(* IEC 61131-3 sources: 2026_Projet_YGO_ExcavatriceDragage/CODE/J_SUPERVISION (part 3) *)

(* ---- FB_TroubleshootingView.st ---- *)
(* ═══════════════════════════════════════════════════════════════
   🕵️♂️ FB_TroubleshootingView — Mise en forme lecture seule pour dépannage
   ───────────────────────────────────────────────────────────────
   📄 Doc : DOC/AF/AF_Partie-14_Fonction_Troubleshooting/FB_TroubleshootingView_v1.2.md
   🔗 Producteur unique de GVL_Troubleshooting.* — instancié UNE SEULE FOIS,
      dans PRG_07_Supervision, après §3 Projections IHM.
   🔒 Lecture seule stricte : aucune VAR_OUTPUT de commande, aucun calcul métier,
      aucune fusion de source — pure recopie de faits déjà publiés ailleurs.
   ⚠️ WinchM2 est typé ST_WinchBenneHMI (pas ST_WinchHMI comme WinchM1) : ce lot
      (LOT_TROUBLESHOOTING_VIEW_ET_WINCHHMI) a introduit ST_WinchBenneHMI pour porter
      Bucket côté M2 uniquement (GVL_IHM.M2TreuilBenne) — adaptation du port fiche §3
      nécessaire suite à AC5 (Bucket retiré de ST_WinchHMI commun M1/M2).
   Écriture GVL directe : seule exception au principe "pas de GVL comme bus de
      commande" (AF_Partie-03 §5) — GVL_Troubleshooting n'est jamais relue par un FB
      métier, uniquement par Watch CODESYS / export SCADA dépannage (fiche §3/§7).
   ⚠️ Idx201_JoystickSelected (ContexteMachineGlobal) lit GVL_IHM.Modes.Cmd.TglJoystickMaster
      directement (variable globale IEC 61131-3, visible sans passage par VAR_INPUT) — ce
      port n'est pas dans la table fiche §3 mais le producteur exact est documenté fiche §5.1.
   ═══════════════════════════════════════════════════════════════ *)
FUNCTION_BLOCK PUBLIC FB_TroubleshootingView
VAR_INPUT
    Enable                   : BOOL; (* --> [CMD] TRUE en permanence — fiche §3, aucune condition de scan *)

    (* 📡 PRG_02_Acquisition *)
    HwIn                     : ST_HardwareImage;   (* --> [HW] Image entrées qualifiées *)
    HwReal                   : ST_HardwareImage;   (* --> [HW] Image entrées réelles *)
    InputModuleFault         : BOOL;   (* --> [HW] Défaut module d'entrée *)
    LocalDigitalIoOk         : BOOL; (* --> [HW] Mirroir Network.InputModules — pas de champ ST_Chain* dédié ce lot *)
    Vh0800EndOk              : BOOL; (* --> [HW] idem *)
    Vh0808EtpOk              : BOOL; (* --> [HW] idem *)

    (* 🎚️ PRG_03_Modes_Cycle *)
    Auth                     : ST_Modes_Autorisations;   (* --> [SAFE] Autorisations machine *)

    (* 🛗 PRG_04_Treuils_Benne — demandes publiques déjà arbitrées *)
    M1LogicRequestSpeedCmd_Pct : REAL;   (* --> [CMD] Consigne vitesse M1 *)
    M1LogicRequestDirection    : INT;   (* --> [CMD] Sens M1 *)
    M2LogicRequestSpeedCmd_Pct : REAL;   (* --> [CMD] Consigne vitesse M2 *)
    M2LogicRequestDirection    : INT;   (* --> [CMD] Sens M2 *)
    WinchBothMotionDirection : INT;   (* --> [CMD] Direction couplée *)
    WinchBothMotionActive    : BOOL;   (* --> [CMD] Demande couplée active *)
    CycleAutoBusy                : BOOL;   (* --> [HW] Cycle auto actif *)
    CycleM1SpeedTgt_Pct          : REAL;   (* --> [CMD] Consigne cycle M1 *)
    CycleM2SpeedTgt_Pct          : REAL;   (* --> [CMD] Consigne cycle M2 *)
    CycleBucketOpen              : BOOL;   (* --> [HW] Benne ouverte cycle *)
    CycleTargetPosition          : INT;   (* --> [CMD] Cible cycle *)

    (* 🎭 GVL_Simulation *)
    SimulationModeActive     : BOOL;   (* --> [TST] Mode simulation *)
    SimWinchActive           : BOOL;   (* --> [TST] Sim treuils *)
    SimTranslationActive     : BOOL;   (* --> [TST] Sim translation *)
    SimOperatorActive        : BOOL;   (* --> [TST] Sim opérateur *)
    SimSafetyActive          : BOOL;   (* --> [TST] Sim sécurité *)

    (* 🛗 GVL_IHM — images publiques déjà produites *)
    WinchM1                  : ST_WinchHMI;      (* --> [HW] GVL_IHM.M1TreuilRetenue *)
    WinchM2                  : ST_WinchBenneHMI; (* --> [HW] GVL_IHM.M2TreuilBenne — porte Bucket *)
    Sync                     : ST_SyncHMI;       (* --> [HW] GVL_IHM.M1M2Sync *)
    Translation              : ST_TranslationHMI;(* --> [HW] GVL_IHM.M3Translation *)
    Commun                   : ST_CommunHMI;     (* --> [HW] GVL_IHM.Commun *)
    Network                  : ST_NetworkDiagHMI;(* --> [HW] GVL_IHM.Network *)
    JoystickHMI              : ST_JoystickHMI;   (* --> [HW] GVL_IHM.JOY1Joystick *)
    Permits                  : ST_PermitVisibilityHMI; (* --> [DIAG] Vue unique des permis produite par PRG_07 *)

    (* 🛡️ Sorties publiques AU produites par PRG_06_Outputs *)
    EmergencyState           : ST_Safety_Emergency_State;   (* --> [SAFE] État AU *)
    EmergencyDiag            : ST_Safety_Emergency_Diag;   (* --> [SAFE] Diagnostic AU *)
    PowerCutOffActive        : BOOL;   (* --> [SAFE] Coupure puissance *)
    ArmingPulseActive        : BOOL;   (* --> [SAFE] Impulsion réarmement *)
    MaintainAActive          : BOOL;   (* --> [SAFE] Maintien canal A *)
    MaintainBActive          : BOOL;   (* --> [SAFE] Maintien canal B *)

    (* 📤 Ordres finaux produits par PRG_06_Outputs, après barrière et protecteurs *)
    Outputs                  : ST_OutputsInterPrg; (* --> [CMD] Ordres actionneurs finaux *)
    CmdM3DriveFreqWord       : WORD;   (* --> [CMD] Consigne finale variateur M3 [0.01 Hz] *)

    (* 🔄 Séquenceur de cycle semi-automatique *)
    CycleReady               : BOOL;   (* --> [STAT] Séquenceur prêt *)
    CycleDone                : BOOL;   (* --> [STAT] Séquenceur terminé *)
    CycleError               : BOOL;   (* --> [STAT] Séquenceur en erreur *)
    CycleErrorId             : WORD;   (* --> [DIAG] Code erreur séquenceur *)
    CycleFaultLatched        : BOOL;   (* --> [STAT] Défaut latché séquenceur (bloque AX0->AX1, exige Reset) *)
    CycleFaultLatchedId      : WORD;   (* --> [DIAG] Bitfield défaut latché figé *)
    CycleChecksInhibited     : BOOL;   (* --> [TST] Contrôles procédé inhibés *)
    CycleIgnoredCheckId      : WORD;   (* --> [DIAG] Contrôles procédé ignorés *)
    CycleForceStepResult     : STRING(120); (* --> [DIAG] Motif de rejet de la consigne de forcage de step (T358) *)
    CycleStep                : E_AutoCycleStep; (* --> [STAT] Étape courante *)
    CycleStepStr             : STRING(80);  (* --> [STAT] Libellé étape *)
    CycleStepAtError         : E_AutoCycleStep; (* --> [DIAG] Étape au défaut *)
    CycleWaitingForOperator  : BOOL;        (* --> [STAT] Attente action humaine *)
    CycleWaitingForProcess   : BOOL;        (* --> [STAT] Attente condition procédé *)
    CycleOperatorActionId    : WORD;        (* --> [DIAG] ID action attendue *)
    CycleOperatorAction      : STRING(120); (* --> [DIAG] Consigne explicite *)
    CycleExpectedAxis        : E_OperatorAxis; (* --> [STAT] Organe attendu *)
    CycleExpectedDirection   : INT;         (* --> [STAT] Sens attendu (-1, 0, +1) *)
    CycleStartRequest        : BOOL;   (* --> [CMD] Demande Start *)
    CycleAbortRequest        : BOOL;   (* --> [CMD] Demande Abort *)
    CycleTargetDepth_M       : REAL;   (* --> [CFG] Profondeur consigne *)
    CycleKoboldBottomTouch   : BOOL;   (* --> [HW] Contact fond *)
    CycleSpeedMismatchActive : BOOL;   (* --> [DIAG] Écart vitesse M1/M2 *)
    CycleLimitLegalReached   : BOOL;   (* --> [SAFE] Limite légale atteinte *)
    CycleWinchSyncError      : BOOL;   (* --> [SAFE] Erreur synchro treuils *)
    CycleM1SpeedStepApplied  : INT;    (* --> [HW] Palier vitesse appliqué M1 (0..5, causes 8/9 FB_CycleSemiAuto) *)
    CycleM2SpeedStepApplied  : INT;    (* --> [HW] Palier vitesse appliqué M2 (0..5, causes 8/9 FB_CycleSemiAuto) *)
    CycleAutoDiveM2Step5Active : BOOL; (* --> [STAT] Essai T291-A actif (M2 cible palier 5 en plongée) *)
    CycleM1SpeedStepAtFault  : INT;    (* --> [DIAG] Palier M1 appliqué, figé au moment du défaut (0..5) *)
    CycleM2SpeedStepAtFault  : INT;    (* --> [DIAG] Palier M2 appliqué, figé au moment du défaut (0..5) *)
    JoystickDeadmanArmed     : BOOL;   (* --> [CMD] Homme-mort armé *)
    JoystickAtNeutral        : BOOL;   (* --> [HW] Joystick au neutre *)
    HomedM1                  : BOOL;   (* --> [HW] Codeur M1 référencé *)
    HomedM2                  : BOOL;   (* --> [HW] Codeur M2 référencé *)

    (* 📐 Config effective limite haute — source _CommunCfgPersist (≠ copie IHM) *)
    CfgTopLimitM             : REAL;   (* --> [CFG] Limite haute active (m) = CfgCableLimitAscent_M *)

    (* 🕵️ PRG_04/05 — Trace de blocage terrain (cause priorisée + horodatage, produite
       par PRG_04 §8bis / PRG_05 §4bis, publiée via Data ; pure recopie ici) *)
    WinchM1Trace             : ST_TraceWinch;       (* --> [DIAG] Trace blocage treuil M1 *)
    WinchM2Trace             : ST_TraceWinch;       (* --> [DIAG] Trace blocage treuil M2 *)
    TranslationTrace         : ST_TraceTranslation; (* --> [DIAG] Trace blocage translation M3 *)
    MachineHoming            : ST_MachineHoming;    (* --> [DIAG] Etat public du cycle de homing conjoint *)
END_VAR
VAR_OUTPUT
    Ready                    : BOOL; (* <-- [STAT] Diagnostic interne minimal — fiche §3 *)
END_VAR

// 🛑 GATE — neutralisation ; aucune écriture GVL_Troubleshooting si Enable=FALSE
IF NOT Enable THEN
    Ready := FALSE;
    RETURN;
END_IF;
Ready := TRUE;

{region "§0 Contexte machine global"}
// === 🌐 0. ContexteMachineGlobal : ST_ChainContextGlobal (fiche §5.1) ===
GVL_Troubleshooting.A_ContexteMachineGlobal.Idx101_ModeActive        := Auth.Mode;
GVL_Troubleshooting.A_ContexteMachineGlobal.Idx102_SimulationEnabled := SimulationModeActive;
GVL_Troubleshooting.A_ContexteMachineGlobal.Idx103_JoystickCommOk    := Network.Joystick.Operational;
GVL_Troubleshooting.A_ContexteMachineGlobal.Idx201_JoystickSelected  := GVL_IHM.Modes.Cmd.TglJoystickMaster;
GVL_Troubleshooting.A_ContexteMachineGlobal.Idx202_BypassNetworkGlobal := Network.Bypass.Global;
GVL_Troubleshooting.A_ContexteMachineGlobal.Idx203_BypassSensorsGlobal := FALSE; // TBD non câblé - voir fiche §6 (agrégat multi-domaine à définir)
GVL_Troubleshooting.A_ContexteMachineGlobal.Idx301_EmergencyChainClosed := HwIn.Machine.EmergencyChainClosed_DI;
GVL_Troubleshooting.A_ContexteMachineGlobal.Idx302_PowerContactorEngaged := HwIn.Machine.PowerContactorEngaged_DI;
// Agrégat simple OR de faits déjà publiés (fiche §5.1) — pas un nouveau calcul métier
GVL_Troubleshooting.A_ContexteMachineGlobal.Idx303_SafeStopActiveAny := WinchM1.Safety.SafeStop OR WinchM2.Safety.SafeStop OR Translation.Safety.SafeStop;
GVL_Troubleshooting.A_ContexteMachineGlobal.Idx304_PowerCutOffActiveAny := WinchM1.Safety.PowerCutOff OR WinchM2.Safety.PowerCutOff OR Translation.Safety.PowerCutOff;
GVL_Troubleshooting.A_ContexteMachineGlobal.Idx401_HmiHeartbeatOk    := Commun.HeartbeatIhmOk;
GVL_Troubleshooting.A_ContexteMachineGlobal.Idx402_CycleAutoBusy     := CycleAutoBusy;

{endregion}

{region "§1 Levage synchronise M1/M2"}
// === 🛗 1. LevageSynchroniseM1M2 : ST_ChainWinchSync (fiche §5.2) ===
GVL_Troubleshooting.H_LevageSynchroniseM1M2.Idx101_M1_CablePos_M  := WinchM1.State.Position_M;
GVL_Troubleshooting.H_LevageSynchroniseM1M2.Idx102_M2_CablePos_M  := WinchM2.State.Position_M;
GVL_Troubleshooting.H_LevageSynchroniseM1M2.Idx103_SyncDelta_M    := Sync.State.DeltaPos_M;
GVL_Troubleshooting.H_LevageSynchroniseM1M2.Idx202_SyncEnabled_IHM := Sync.Cmd.SelSyncEnable;
GVL_Troubleshooting.H_LevageSynchroniseM1M2.Idx301_EmergencyChainClosed := HwIn.Machine.EmergencyChainClosed_DI;
GVL_Troubleshooting.H_LevageSynchroniseM1M2.Idx302_SyncFaultActive := Sync.State.Error;
GVL_Troubleshooting.H_LevageSynchroniseM1M2.Idx303_M1_AscentPermit := WinchM1.Safety.AscentPermit;
GVL_Troubleshooting.H_LevageSynchroniseM1M2.Idx304_M2_AscentPermit := WinchM2.Safety.AscentPermit;
GVL_Troubleshooting.H_LevageSynchroniseM1M2.Idx501_M1_CmdRelayFwd_DQ := Outputs.M1RelayFwd;
GVL_Troubleshooting.H_LevageSynchroniseM1M2.Idx502_M2_CmdRelayFwd_DQ := Outputs.M2RelayFwd;
// Idx201_JoyYRaw_Pct / Idx203_ArbitratedSpeed_Pct / Idx303-304_AscentPermit / Idx401_SyncMotionAllowed /
// Idx402-403_SetpointSpeed : non câblés — fiche §5.2 "(reste) champs à revoir un par un", laissés à
// leur valeur d'initialisation, pas de calcul inventé (fiche §7).

{endregion}

{region "§2 Levage unitaire M1/M2"}
// === 🛗 2. LevageUnitaireM1 / LevageUnitaireM2 : ST_ChainWinch (fiche §5.3) ===
// --- M1 ---
GVL_Troubleshooting.I_LevageUnitaireM1.Inputs_100.Idx101_EncoderRawPos := UDINT_TO_DINT(HwIn.Winch.COD1_PosValue);
GVL_Troubleshooting.I_LevageUnitaireM1.Inputs_100.Idx102_CablePos_M := WinchM1.State.Position_M;
GVL_Troubleshooting.I_LevageUnitaireM1.Inputs_100.Idx103_ContactorsReleased_DI := HwIn.Winch.M1_ContactorsReleased_DI;
GVL_Troubleshooting.I_LevageUnitaireM1.Inputs_100.Idx104_BrakeApplied := NOT HwIn.Winch.M1_BrakeIsOpen_DI;
GVL_Troubleshooting.I_LevageUnitaireM1.Inputs_100.Idx105_ThermalOk_DI := HwIn.Winch.M1_ThermalOk_DI;

GVL_Troubleshooting.I_LevageUnitaireM1.Demandes_200.Idx201_JoyRawPhysical_ANA := HwIn.Operator.JoyYRaw_ANA2;
GVL_Troubleshooting.I_LevageUnitaireM1.Demandes_200.Idx202_JoyScaledPhysical_Pct := JoystickHMI.State.AxisCmdY.Deflection;
GVL_Troubleshooting.I_LevageUnitaireM1.Demandes_200.Idx203_HmiManualCmd_BtnAscent := WinchM1.Cmd.BtnAscent;
GVL_Troubleshooting.I_LevageUnitaireM1.Demandes_200.Idx204_HmiManualCmd_BtnDescent := WinchM1.Cmd.BtnDescent;
GVL_Troubleshooting.I_LevageUnitaireM1.Demandes_200.Idx205_CycleAutoCmd_Pct := CycleM1SpeedTgt_Pct;
GVL_Troubleshooting.I_LevageUnitaireM1.Demandes_200.Idx206_ModeActive := Auth.Mode;
GVL_Troubleshooting.I_LevageUnitaireM1.Demandes_200.Idx207_BypassOperatorComm := WinchM1.Bypass.OperatorComm;
GVL_Troubleshooting.I_LevageUnitaireM1.Demandes_200.Idx208_ArbitratedSpeed_Pct := M1LogicRequestSpeedCmd_Pct;
GVL_Troubleshooting.I_LevageUnitaireM1.Demandes_200.Idx209_ArbitratedDirection := M1LogicRequestDirection;
GVL_Troubleshooting.I_LevageUnitaireM1.Demandes_200.Idx210_CoupledUserRequestDirection := WinchBothMotionDirection;
GVL_Troubleshooting.I_LevageUnitaireM1.Demandes_200.Idx211_CoupledUserRequestActive := WinchBothMotionActive;

GVL_Troubleshooting.I_LevageUnitaireM1.Safety_300.Idx301_EmergencyChainClosed := HwIn.Machine.EmergencyChainClosed_DI;
GVL_Troubleshooting.I_LevageUnitaireM1.Safety_300.Idx302_SafeStopActive := WinchM1.Safety.SafeStop;
GVL_Troubleshooting.I_LevageUnitaireM1.Safety_300.Idx303_PowerCutOffActive := WinchM1.Safety.PowerCutOff;
GVL_Troubleshooting.I_LevageUnitaireM1.Safety_300.Idx304_TopSensorPhysical_DI := HwIn.Winch.M1M2_TopPositionFree_DI;
GVL_Troubleshooting.I_LevageUnitaireM1.Safety_300.Idx305_TopSensorBypassActive := Commun.SimTopSensorBypassActive;
GVL_Troubleshooting.I_LevageUnitaireM1.Safety_300.Idx306_AscentPermitEffective := WinchM1.Safety.AscentPermit;
GVL_Troubleshooting.I_LevageUnitaireM1.Safety_300.Idx307_SlackCablePhysical_DI := NOT HwIn.Winch.M2_TensionedCable_DI; // Capteur unique partagé, même signal que SlackCableDetected M1
GVL_Troubleshooting.I_LevageUnitaireM1.Safety_300.Idx308_SlackCableBypassActive := Commun.SimSlackCableBypassActive;
GVL_Troubleshooting.I_LevageUnitaireM1.Safety_300.Idx309_DescendPermitEffective := WinchM1.Safety.DescendPermit;
GVL_Troubleshooting.I_LevageUnitaireM1.Safety_300.Idx310_ErrorOperatorComm := WinchM1.Safety.ErrorOperatorComm;
GVL_Troubleshooting.I_LevageUnitaireM1.Safety_300.Idx311_ErrorEncoder      := WinchM1.Safety.ErrorEncoder;
GVL_Troubleshooting.I_LevageUnitaireM1.Safety_300.Idx312_ErrorPhaseRotation:= WinchM1.Safety.ErrorPhaseRotation;
GVL_Troubleshooting.I_LevageUnitaireM1.Safety_300.Idx313_ErrorMecaA        := WinchM1.Safety.ErrorMecaA;
GVL_Troubleshooting.I_LevageUnitaireM1.Safety_300.Idx314_ErrorMecaB        := WinchM1.Safety.ErrorMecaB;
GVL_Troubleshooting.I_LevageUnitaireM1.Safety_300.Idx315_ErrorMecaC        := WinchM1.Safety.ErrorMecaC;
GVL_Troubleshooting.I_LevageUnitaireM1.Safety_300.Idx316_ErrorMecaD        := WinchM1.Safety.ErrorMecaD;
GVL_Troubleshooting.I_LevageUnitaireM1.Safety_300.Idx317_ErrorMecaE        := WinchM1.Safety.ErrorMecaE;
GVL_Troubleshooting.I_LevageUnitaireM1.Safety_300.Idx318_ErrorBrakeThermal := WinchM1.Safety.ErrorBrakeThermal;
GVL_Troubleshooting.I_LevageUnitaireM1.Safety_300.Idx319_ErrorOppositeDir  := WinchM1.Safety.ErrorOppositeDir;
GVL_Troubleshooting.I_LevageUnitaireM1.Safety_300.Idx320_ErrorNoMovement   := WinchM1.Safety.ErrorNoMovement;
// ⛔ Bloc "limite haute" — pourquoi la montée ne s'arrête pas (M1)
GVL_Troubleshooting.I_LevageUnitaireM1.Safety_300.Idx321_CfgTopLimitM               := CfgTopLimitM;
GVL_Troubleshooting.I_LevageUnitaireM1.Safety_300.Idx322_CablePosM                  := WinchM1.State.Position_M;
GVL_Troubleshooting.I_LevageUnitaireM1.Safety_300.Idx323_TopLimitReached            := WinchM1.Safety.CableLimitAscent;
GVL_Troubleshooting.I_LevageUnitaireM1.Safety_300.Idx324_AscentBlockedByTopLimit    := WinchM1.Safety.CableLimitAscent AND NOT (WinchM1.Bypass.TopLimitSoftware OR Commun.Bypass.TopLimitSoftware);
GVL_Troubleshooting.I_LevageUnitaireM1.Safety_300.Idx325_BypassTopLimitSoftware     := WinchM1.Bypass.TopLimitSoftware;
GVL_Troubleshooting.I_LevageUnitaireM1.Safety_300.Idx326_BypassTopLimitSoftCommun   := Commun.Bypass.TopLimitSoftware;
GVL_Troubleshooting.I_LevageUnitaireM1.Safety_300.Idx327_BypassTopLimitSwitch       := WinchM1.Bypass.TopLimitSwitch;
GVL_Troubleshooting.I_LevageUnitaireM1.Safety_300.Idx328_BypassTopLimitSwitchCommun := Commun.Bypass.TopLimitSwitch;
GVL_Troubleshooting.I_LevageUnitaireM1.Safety_300.Idx329_BypassGlobal               := WinchM1.Bypass.Global;
GVL_Troubleshooting.I_LevageUnitaireM1.Safety_300.Idx330_BypassGlobalCommun         := Commun.Bypass.Global;

GVL_Troubleshooting.I_LevageUnitaireM1.Control_400.Idx401_MotionAllowed := WinchM1.State.Ready;
GVL_Troubleshooting.I_LevageUnitaireM1.Control_400.Idx402_SpeedStepCalculated := WinchM1.State.StepNumber;
GVL_Troubleshooting.I_LevageUnitaireM1.Control_400.Idx403_SpeedRamp_Pct := WinchM1.State.SpeedCmd_Pct;
GVL_Troubleshooting.I_LevageUnitaireM1.Control_400.Idx404_BrakeReleaseAuthorized := WinchM1.State.BrakeCmd;
GVL_Troubleshooting.I_LevageUnitaireM1.Control_400.Idx405_FinalInterlockState := WinchM1.State.FinalInterlockState;
GVL_Troubleshooting.I_LevageUnitaireM1.Control_400.Idx406_FinalInterlockReason := WinchM1.State.FinalInterlockReason;
GVL_Troubleshooting.I_LevageUnitaireM1.Control_400.Idx407_FinalAuthorizedStep := WinchM1.State.FinalAuthorizedStep;
GVL_Troubleshooting.I_LevageUnitaireM1.Control_400.Idx408_BrakeCommandOpenConfirmed := WinchM1.State.BrakeCommandOpenConfirmed;
GVL_Troubleshooting.I_LevageUnitaireM1.Control_400.Idx409_BrakeTimeoutElapsed := WinchM1.State.FinalBrakeTimeoutElapsed;
GVL_Troubleshooting.I_LevageUnitaireM1.Control_400.Idx410_RestartDelayElapsed := WinchM1.State.FinalRestartDelayElapsed;
GVL_Troubleshooting.I_LevageUnitaireM1.Control_400.Idx411_StepDelayElapsed := WinchM1.State.FinalStepDelayElapsed;
GVL_Troubleshooting.I_LevageUnitaireM1.Control_400.Idx412_InTopSlowdownZone := WinchM1.State.InTopSlowdownZone;
GVL_Troubleshooting.I_LevageUnitaireM1.Control_400.Idx413_InBottomSlowdownZone := WinchM1.State.InBottomSlowdownZone;
GVL_Troubleshooting.I_LevageUnitaireM1.Control_400.Idx414_BottomLimitActiveM := WinchM1.State.BottomLimitActiveM;
GVL_Troubleshooting.I_LevageUnitaireM1.Control_400.Idx415_MotorRequest := WinchM1.State.FinalMotorRequest;
GVL_Troubleshooting.I_LevageUnitaireM1.Control_400.Idx416_RestartRequired := WinchM1.State.FinalRestartRequired;
GVL_Troubleshooting.I_LevageUnitaireM1.Control_400.Idx417_RestartInhibit := WinchM1.State.FinalRestartInhibit;
GVL_Troubleshooting.I_LevageUnitaireM1.Control_400.Idx418_NeutralRequestSeen := WinchM1.State.FinalNeutralRequestSeen;

GVL_Troubleshooting.I_LevageUnitaireM1.Outputs_500.Idx501_CmdRelayAscent_RQ := Outputs.M1RelayFwd;
GVL_Troubleshooting.I_LevageUnitaireM1.Outputs_500.Idx502_CmdRelayDescent_RQ := Outputs.M1RelayRev;
GVL_Troubleshooting.I_LevageUnitaireM1.Outputs_500.Idx503_CmdSpeedContactor1_DQ := Outputs.M1SpeedContactor1;
GVL_Troubleshooting.I_LevageUnitaireM1.Outputs_500.Idx504_CmdSpeedContactor4_DQ := Outputs.M1SpeedContactor4;
GVL_Troubleshooting.I_LevageUnitaireM1.Outputs_500.Idx505_CmdBrakeRelease_RQ := WinchM1.State.BrakeCmd;

// --- M2 (même patron, source WinchM2) ---
GVL_Troubleshooting.J_LevageUnitaireM2.Inputs_100.Idx101_EncoderRawPos := UDINT_TO_DINT(HwIn.Winch.COD2_PosValue);
GVL_Troubleshooting.J_LevageUnitaireM2.Inputs_100.Idx102_CablePos_M := WinchM2.State.Position_M;
GVL_Troubleshooting.J_LevageUnitaireM2.Inputs_100.Idx103_ContactorsReleased_DI := HwIn.Winch.M2_ContactorsReleased_DI;
GVL_Troubleshooting.J_LevageUnitaireM2.Inputs_100.Idx104_BrakeApplied := NOT HwIn.Winch.M2_BrakeIsOpen_DI;
GVL_Troubleshooting.J_LevageUnitaireM2.Inputs_100.Idx105_ThermalOk_DI := HwIn.Winch.M2_ThermalOk_DI;

GVL_Troubleshooting.J_LevageUnitaireM2.Demandes_200.Idx201_JoyRawPhysical_ANA := HwIn.Operator.JoyYRaw_ANA2;
GVL_Troubleshooting.J_LevageUnitaireM2.Demandes_200.Idx202_JoyScaledPhysical_Pct := JoystickHMI.State.AxisCmdY.Deflection;
GVL_Troubleshooting.J_LevageUnitaireM2.Demandes_200.Idx203_HmiManualCmd_BtnAscent := WinchM2.Cmd.BtnAscent;
GVL_Troubleshooting.J_LevageUnitaireM2.Demandes_200.Idx204_HmiManualCmd_BtnDescent := WinchM2.Cmd.BtnDescent;
GVL_Troubleshooting.J_LevageUnitaireM2.Demandes_200.Idx205_CycleAutoCmd_Pct := CycleM2SpeedTgt_Pct;
GVL_Troubleshooting.J_LevageUnitaireM2.Demandes_200.Idx206_ModeActive := Auth.Mode;
GVL_Troubleshooting.J_LevageUnitaireM2.Demandes_200.Idx207_BypassOperatorComm := WinchM2.Bypass.OperatorComm;
GVL_Troubleshooting.J_LevageUnitaireM2.Demandes_200.Idx208_ArbitratedSpeed_Pct := M2LogicRequestSpeedCmd_Pct;
GVL_Troubleshooting.J_LevageUnitaireM2.Demandes_200.Idx209_ArbitratedDirection := M2LogicRequestDirection;
GVL_Troubleshooting.J_LevageUnitaireM2.Demandes_200.Idx210_CoupledUserRequestDirection := WinchBothMotionDirection;
GVL_Troubleshooting.J_LevageUnitaireM2.Demandes_200.Idx211_CoupledUserRequestActive := WinchBothMotionActive;

GVL_Troubleshooting.J_LevageUnitaireM2.Safety_300.Idx301_EmergencyChainClosed := HwIn.Machine.EmergencyChainClosed_DI;
GVL_Troubleshooting.J_LevageUnitaireM2.Safety_300.Idx302_SafeStopActive := WinchM2.Safety.SafeStop;
GVL_Troubleshooting.J_LevageUnitaireM2.Safety_300.Idx303_PowerCutOffActive := WinchM2.Safety.PowerCutOff;
GVL_Troubleshooting.J_LevageUnitaireM2.Safety_300.Idx304_TopSensorPhysical_DI := HwIn.Winch.M1M2_TopPositionFree_DI;
GVL_Troubleshooting.J_LevageUnitaireM2.Safety_300.Idx305_TopSensorBypassActive := Commun.SimTopSensorBypassActive;
GVL_Troubleshooting.J_LevageUnitaireM2.Safety_300.Idx306_AscentPermitEffective := WinchM2.Safety.AscentPermit;
// Bug affichage MES 2026-09-04 : publiait TensionedCable_DI sans l'inverser -> cable
// tendu (bon) s'affichait comme "mou detecte". Logique securite reelle (PRG_04) deja
// correcte (NOT TensionedCable_DI) ; seul ce mirroir troubleshooting etait faux.
GVL_Troubleshooting.J_LevageUnitaireM2.Safety_300.Idx307_SlackCablePhysical_DI := NOT HwIn.Winch.M2_TensionedCable_DI;
GVL_Troubleshooting.J_LevageUnitaireM2.Safety_300.Idx308_SlackCableBypassActive := Commun.SimSlackCableBypassActive;
GVL_Troubleshooting.J_LevageUnitaireM2.Safety_300.Idx309_DescendPermitEffective := WinchM2.Safety.DescendPermit;
GVL_Troubleshooting.J_LevageUnitaireM2.Safety_300.Idx310_ErrorOperatorComm := WinchM2.Safety.ErrorOperatorComm;
GVL_Troubleshooting.J_LevageUnitaireM2.Safety_300.Idx311_ErrorEncoder      := WinchM2.Safety.ErrorEncoder;
GVL_Troubleshooting.J_LevageUnitaireM2.Safety_300.Idx312_ErrorPhaseRotation:= WinchM2.Safety.ErrorPhaseRotation;
GVL_Troubleshooting.J_LevageUnitaireM2.Safety_300.Idx313_ErrorMecaA        := WinchM2.Safety.ErrorMecaA;
GVL_Troubleshooting.J_LevageUnitaireM2.Safety_300.Idx314_ErrorMecaB        := WinchM2.Safety.ErrorMecaB;
GVL_Troubleshooting.J_LevageUnitaireM2.Safety_300.Idx315_ErrorMecaC        := WinchM2.Safety.ErrorMecaC;
GVL_Troubleshooting.J_LevageUnitaireM2.Safety_300.Idx316_ErrorMecaD        := WinchM2.Safety.ErrorMecaD;
GVL_Troubleshooting.J_LevageUnitaireM2.Safety_300.Idx317_ErrorMecaE        := WinchM2.Safety.ErrorMecaE;
GVL_Troubleshooting.J_LevageUnitaireM2.Safety_300.Idx318_ErrorBrakeThermal := WinchM2.Safety.ErrorBrakeThermal;
GVL_Troubleshooting.J_LevageUnitaireM2.Safety_300.Idx319_ErrorOppositeDir  := WinchM2.Safety.ErrorOppositeDir;
GVL_Troubleshooting.J_LevageUnitaireM2.Safety_300.Idx320_ErrorNoMovement   := WinchM2.Safety.ErrorNoMovement;
// ⛔ Bloc "limite haute" — pourquoi la montée ne s'arrête pas (M2, sans M2_LimitShift ici)
GVL_Troubleshooting.J_LevageUnitaireM2.Safety_300.Idx321_CfgTopLimitM               := CfgTopLimitM;
GVL_Troubleshooting.J_LevageUnitaireM2.Safety_300.Idx322_CablePosM                  := WinchM2.State.Position_M;
GVL_Troubleshooting.J_LevageUnitaireM2.Safety_300.Idx323_TopLimitReached            := WinchM2.Safety.CableLimitAscent;
GVL_Troubleshooting.J_LevageUnitaireM2.Safety_300.Idx324_AscentBlockedByTopLimit    := WinchM2.Safety.CableLimitAscent AND NOT (WinchM2.Bypass.TopLimitSoftware OR Commun.Bypass.TopLimitSoftware);
GVL_Troubleshooting.J_LevageUnitaireM2.Safety_300.Idx325_BypassTopLimitSoftware     := WinchM2.Bypass.TopLimitSoftware;
GVL_Troubleshooting.J_LevageUnitaireM2.Safety_300.Idx326_BypassTopLimitSoftCommun   := Commun.Bypass.TopLimitSoftware;
GVL_Troubleshooting.J_LevageUnitaireM2.Safety_300.Idx327_BypassTopLimitSwitch       := WinchM2.Bypass.TopLimitSwitch;
GVL_Troubleshooting.J_LevageUnitaireM2.Safety_300.Idx328_BypassTopLimitSwitchCommun := Commun.Bypass.TopLimitSwitch;
GVL_Troubleshooting.J_LevageUnitaireM2.Safety_300.Idx329_BypassGlobal               := WinchM2.Bypass.Global;
GVL_Troubleshooting.J_LevageUnitaireM2.Safety_300.Idx330_BypassGlobalCommun         := Commun.Bypass.Global;

GVL_Troubleshooting.J_LevageUnitaireM2.Control_400.Idx401_MotionAllowed := WinchM2.State.Ready;
GVL_Troubleshooting.J_LevageUnitaireM2.Control_400.Idx402_SpeedStepCalculated := WinchM2.State.StepNumber;
GVL_Troubleshooting.J_LevageUnitaireM2.Control_400.Idx403_SpeedRamp_Pct := WinchM2.State.SpeedCmd_Pct;
GVL_Troubleshooting.J_LevageUnitaireM2.Control_400.Idx404_BrakeReleaseAuthorized := WinchM2.State.BrakeCmd;
GVL_Troubleshooting.J_LevageUnitaireM2.Control_400.Idx405_FinalInterlockState := WinchM2.State.FinalInterlockState;
GVL_Troubleshooting.J_LevageUnitaireM2.Control_400.Idx406_FinalInterlockReason := WinchM2.State.FinalInterlockReason;
GVL_Troubleshooting.J_LevageUnitaireM2.Control_400.Idx407_FinalAuthorizedStep := WinchM2.State.FinalAuthorizedStep;
GVL_Troubleshooting.J_LevageUnitaireM2.Control_400.Idx408_BrakeCommandOpenConfirmed := WinchM2.State.BrakeCommandOpenConfirmed;
GVL_Troubleshooting.J_LevageUnitaireM2.Control_400.Idx409_BrakeTimeoutElapsed := WinchM2.State.FinalBrakeTimeoutElapsed;
GVL_Troubleshooting.J_LevageUnitaireM2.Control_400.Idx410_RestartDelayElapsed := WinchM2.State.FinalRestartDelayElapsed;
GVL_Troubleshooting.J_LevageUnitaireM2.Control_400.Idx411_StepDelayElapsed := WinchM2.State.FinalStepDelayElapsed;
GVL_Troubleshooting.J_LevageUnitaireM2.Control_400.Idx412_InTopSlowdownZone := WinchM2.State.InTopSlowdownZone;
GVL_Troubleshooting.J_LevageUnitaireM2.Control_400.Idx413_InBottomSlowdownZone := WinchM2.State.InBottomSlowdownZone;
GVL_Troubleshooting.J_LevageUnitaireM2.Control_400.Idx414_BottomLimitActiveM := WinchM2.State.BottomLimitActiveM;
GVL_Troubleshooting.J_LevageUnitaireM2.Control_400.Idx415_MotorRequest := WinchM2.State.FinalMotorRequest;
GVL_Troubleshooting.J_LevageUnitaireM2.Control_400.Idx416_RestartRequired := WinchM2.State.FinalRestartRequired;
GVL_Troubleshooting.J_LevageUnitaireM2.Control_400.Idx417_RestartInhibit := WinchM2.State.FinalRestartInhibit;
GVL_Troubleshooting.J_LevageUnitaireM2.Control_400.Idx418_NeutralRequestSeen := WinchM2.State.FinalNeutralRequestSeen;

GVL_Troubleshooting.J_LevageUnitaireM2.Outputs_500.Idx501_CmdRelayAscent_RQ := Outputs.M2RelayFwd;
GVL_Troubleshooting.J_LevageUnitaireM2.Outputs_500.Idx502_CmdRelayDescent_RQ := Outputs.M2RelayRev;
GVL_Troubleshooting.J_LevageUnitaireM2.Outputs_500.Idx503_CmdSpeedContactor1_DQ := Outputs.M2SpeedContactor1;
GVL_Troubleshooting.J_LevageUnitaireM2.Outputs_500.Idx504_CmdSpeedContactor4_DQ := Outputs.M2SpeedContactor4;
GVL_Troubleshooting.J_LevageUnitaireM2.Outputs_500.Idx505_CmdBrakeRelease_RQ := WinchM2.State.BrakeCmd;

{endregion}

{region "§3 Benne ouverture et fermeture"}
// === 🪣 3. BenneOuvertureFermeture : ST_ChainBucket (fiche §5.4, source WinchM2.Bucket) ===
GVL_Troubleshooting.K_BenneOuvertureFermeture.Idx101_BucketIsOpen := WinchM2.Bucket.State.MechState.IsOpen;
GVL_Troubleshooting.K_BenneOuvertureFermeture.Idx102_BucketIsClosed := WinchM2.Bucket.State.MechState.IsClosed;
GVL_Troubleshooting.K_BenneOuvertureFermeture.Idx103_OffsetPos_M := WinchM2.Bucket.State.ActiveOffset_M;
GVL_Troubleshooting.K_BenneOuvertureFermeture.Idx104_AutoSeqActive := WinchM2.Bucket.State.AutoBucketSeqActive;
GVL_Troubleshooting.K_BenneOuvertureFermeture.Idx105_StateIncoherent := WinchM2.Bucket.State.MechState.StateIncoherent;
GVL_Troubleshooting.K_BenneOuvertureFermeture.Idx106_FBState := WinchM2.Bucket.State.FBState;
GVL_Troubleshooting.K_BenneOuvertureFermeture.Idx107_LastPosM2Open_M := WinchM2.Bucket.State.MechState.LastPosM2Open;
GVL_Troubleshooting.K_BenneOuvertureFermeture.Idx108_LastPosM2Close_M := WinchM2.Bucket.State.MechState.LastPosM2Close;
GVL_Troubleshooting.K_BenneOuvertureFermeture.Idx109_BucketTooOpen := WinchM2.Bucket.State.MechState.TooOpen;
GVL_Troubleshooting.K_BenneOuvertureFermeture.Idx110_BucketTooClosed := WinchM2.Bucket.State.MechState.TooClosed;
GVL_Troubleshooting.K_BenneOuvertureFermeture.Idx111_BucketIsIntermediate := WinchM2.Bucket.State.MechState.IsIntermediate;
GVL_Troubleshooting.K_BenneOuvertureFermeture.Idx112_DeltaPosition_M := WinchM2.Bucket.State.DeltaPosition_M;
GVL_Troubleshooting.K_BenneOuvertureFermeture.Idx113_MachineHomed := WinchM2.Bucket.State.MachineHomed;
GVL_Troubleshooting.K_BenneOuvertureFermeture.Idx114_MachineHomingStep := WinchM2.Bucket.State.MachineHomingStep;
GVL_Troubleshooting.K_BenneOuvertureFermeture.Idx115_MachineHomingFailed := WinchM2.Bucket.State.MachineHomingFailed;
GVL_Troubleshooting.K_BenneOuvertureFermeture.Idx116_M1ReferenceMissing := NOT WinchM1.State.Encoder.Homed OR WinchM1.State.Encoder.HomingSuspect;
GVL_Troubleshooting.K_BenneOuvertureFermeture.Idx117_M2ReferenceMissing := NOT WinchM2.State.Encoder.Homed OR WinchM2.State.Encoder.HomingSuspect;
GVL_Troubleshooting.K_BenneOuvertureFermeture.Idx118_BucketOffsetUnknown := NOT WinchM2.Bucket.State.MechState.ActiveOffsetValid;
GVL_Troubleshooting.K_BenneOuvertureFermeture.Idx119_ReferenceTransaction := WinchM2.Bucket.State.MachineHomingActive;
GVL_Troubleshooting.K_BenneOuvertureFermeture.Idx120_MachineHomingLossSafeStop := WinchM2.Bucket.State.MachineHomingLossSafeStop;
GVL_Troubleshooting.K_BenneOuvertureFermeture.Idx201_HmiCmd_BtnOpen := WinchM2.Bucket.Cmd.BtnOpen;
GVL_Troubleshooting.K_BenneOuvertureFermeture.Idx202_HmiCmd_BtnClose := WinchM2.Bucket.Cmd.BtnClose;
GVL_Troubleshooting.K_BenneOuvertureFermeture.Idx203_CycleCmd_Open := CycleBucketOpen;
GVL_Troubleshooting.K_BenneOuvertureFermeture.Idx204_CoupledDiveOpenArmed := WinchM2.Bucket.State.CoupledDiveOpenArmed;
GVL_Troubleshooting.K_BenneOuvertureFermeture.Idx205_CoupledAscentCloseArmed := WinchM2.Bucket.State.CoupledAscentCloseArmed;
GVL_Troubleshooting.K_BenneOuvertureFermeture.Idx206_CloseReqActive := WinchM2.Bucket.State.CloseActive;
GVL_Troubleshooting.K_BenneOuvertureFermeture.Idx207_OpenReqActive := WinchM2.Bucket.State.OpenActive;
GVL_Troubleshooting.K_BenneOuvertureFermeture.Idx208_MotionBlockedByBucket := WinchM2.Bucket.State.CoupledMotionBlockedByBucket;
GVL_Troubleshooting.K_BenneOuvertureFermeture.Idx301_EmergencyChainClosed := HwIn.Machine.EmergencyChainClosed_DI;
GVL_Troubleshooting.K_BenneOuvertureFermeture.Idx302_BucketFaultActive := WinchM2.Bucket.State.Error;
GVL_Troubleshooting.K_BenneOuvertureFermeture.Idx303_KoboldAutoStopEnabled := Commun.Cfg.TglEnableKoboldAutoStopDescent;
GVL_Troubleshooting.K_BenneOuvertureFermeture.Idx304_KoboldImmersionConfirmed := Commun.KoboldImmersionConfirmed;
GVL_Troubleshooting.K_BenneOuvertureFermeture.Idx305_KoboldBottomTouchLatched := Commun.KoboldBottomTouchLatched;
GVL_Troubleshooting.K_BenneOuvertureFermeture.Idx306_ErrorIdRaw := WinchM2.Bucket.State.ErrorId;
GVL_Troubleshooting.K_BenneOuvertureFermeture.Idx307_EffectivePermit_Open := Permits.EffectivePermitBucket_Open;
GVL_Troubleshooting.K_BenneOuvertureFermeture.Idx308_EffectivePermit_Close := Permits.EffectivePermitBucket_Close;
GVL_Troubleshooting.K_BenneOuvertureFermeture.Idx401_BucketBusy := WinchM2.Bucket.State.Busy;
GVL_Troubleshooting.K_BenneOuvertureFermeture.Idx402_BucketDone := WinchM2.Bucket.State.Done;
GVL_Troubleshooting.K_BenneOuvertureFermeture.Idx403_ExtractionControlActive := WinchM2.Bucket.State.ExtractionControlActive;
GVL_Troubleshooting.K_BenneOuvertureFermeture.Idx501_M2_CmdRev_DQ := Outputs.M2RelayRev; // Ouverture benne = relais descente M2

{endregion}

// §4 Assistance dragage retire : GVL_Troubleshooting ne porte plus ce slot (M_Réserve),
// FB_DiveSearch/FB_ExtractionAssist supprimés (legacy, jamais actifs).

{region "§5 Translation pont M3"}
// === ↔️ 4. TranslationPontM3 : ST_ChainTranslation (fiche §5.5, source Translation) ===
GVL_Troubleshooting.L_TranslationPontM3.Inputs_100.Idx101_PosTremie_DI := Translation.State.PositionTremie;
GVL_Troubleshooting.L_TranslationPontM3.Inputs_100.Idx102_PosPV_DI := Translation.State.PositionPV;
GVL_Troubleshooting.L_TranslationPontM3.Inputs_100.Idx103_PosP2_DI := Translation.State.PositionP2;
GVL_Troubleshooting.L_TranslationPontM3.Inputs_100.Idx104_PosP1_DI := Translation.State.PositionP1;
GVL_Troubleshooting.L_TranslationPontM3.Inputs_100.Idx105_PosMaintenance_DI := Translation.State.PositionMaintenance;
GVL_Troubleshooting.L_TranslationPontM3.Inputs_100.Idx106_DriveActualFreq_Hz := Translation.State.DriveActualFreq_Hz;
GVL_Troubleshooting.L_TranslationPontM3.Inputs_100.Idx107_DriveStatusWord := HwIn.Translation.M3_StatusWord;
GVL_Troubleshooting.L_TranslationPontM3.Inputs_100.Idx108_BrakeApplied := NOT Translation.State.BrakeFeedback;
GVL_Troubleshooting.L_TranslationPontM3.Inputs_100.Idx109_DriveThermalOk := Translation.State.DriveThermalOk;

GVL_Troubleshooting.L_TranslationPontM3.Demandes_200.Idx201_JoyXRaw_ANA := HwIn.Operator.JoyXRaw_ANA1;
GVL_Troubleshooting.L_TranslationPontM3.Demandes_200.Idx202_JoyXScaled_Pct := GVL_IHM.JOY1Joystick.State.AxisCmdX.Deflection;
GVL_Troubleshooting.L_TranslationPontM3.Demandes_200.Idx203_HmiCmd_BtnTremie := Translation.Cmd.BtnTremie;
GVL_Troubleshooting.L_TranslationPontM3.Demandes_200.Idx204_HmiCmd_BtnMaintenance := Translation.Cmd.BtnMaintenance;
GVL_Troubleshooting.L_TranslationPontM3.Demandes_200.Idx205_HmiTargetPosition := Translation.Cmd.SelTarget;
GVL_Troubleshooting.L_TranslationPontM3.Demandes_200.Idx206_CycleTargetPosition := CycleTargetPosition;
GVL_Troubleshooting.L_TranslationPontM3.Demandes_200.Idx207_ModeActive := Auth.Mode;
GVL_Troubleshooting.L_TranslationPontM3.Demandes_200.Idx208_BypassNetworkActive := Translation.Bypass.Global;
GVL_Troubleshooting.L_TranslationPontM3.Demandes_200.Idx209_ArbitratedSpeed_Pct := Translation.State.SpeedCmd_Pct;

GVL_Troubleshooting.L_TranslationPontM3.Safety_300.Idx301_EmergencyChainClosed := HwIn.Machine.EmergencyChainClosed_DI;
GVL_Troubleshooting.L_TranslationPontM3.Safety_300.Idx302_SafeStopActive := Translation.Safety.SafeStop;
GVL_Troubleshooting.L_TranslationPontM3.Safety_300.Idx303_PowerCutOffActive := Translation.Safety.PowerCutOff;
GVL_Troubleshooting.L_TranslationPontM3.Safety_300.Idx304_LimitSwitchTremieActive := Translation.State.LimitSwitchTremie;
GVL_Troubleshooting.L_TranslationPontM3.Safety_300.Idx305_LimitSwitchMaintenanceActive := Translation.State.LimitSwitchMaintenance;
GVL_Troubleshooting.L_TranslationPontM3.Safety_300.Idx306_BypassLimitSwitch := Translation.Bypass.LimitSwitch;
GVL_Troubleshooting.L_TranslationPontM3.Safety_300.Idx307_PositionDecoderIncoherent := Translation.State.SensorWordIncoherent;
GVL_Troubleshooting.L_TranslationPontM3.Safety_300.Idx308_HeightInterlockBlocking := Translation.State.HeightInterlockBlocking;
GVL_Troubleshooting.L_TranslationPontM3.Safety_300.Idx309_ErrorOperatorComm := Translation.Safety.ErrorOperatorComm;
GVL_Troubleshooting.L_TranslationPontM3.Safety_300.Idx310_ErrorDriveComm    := Translation.Safety.ErrorDriveComm;
GVL_Troubleshooting.L_TranslationPontM3.Safety_300.Idx311_ErrorPhaseRotation:= Translation.Safety.ErrorPhaseRotation;
GVL_Troubleshooting.L_TranslationPontM3.Safety_300.Idx312_ErrorBrakeThermal := Translation.Safety.ErrorBrakeThermal;
GVL_Troubleshooting.L_TranslationPontM3.Safety_300.Idx313_ErrorMecaB        := Translation.Safety.ErrorMecaB;
GVL_Troubleshooting.L_TranslationPontM3.Safety_300.Idx314_ErrorMecaA        := Translation.Safety.ErrorMecaA;
GVL_Troubleshooting.L_TranslationPontM3.Safety_300.Idx315_ErrorLimitSwitch  := Translation.Safety.ErrorLimitSwitch;
GVL_Troubleshooting.L_TranslationPontM3.Safety_300.Idx316_ErrorSensorIncoherent := Translation.Safety.ErrorSensorIncoherent;
GVL_Troubleshooting.L_TranslationPontM3.Safety_300.Idx317_ErrorId := Translation.Safety.ErrorId; // Masque brut complet (latch cause, source d'arbitrage PowerCutOff)
GVL_Troubleshooting.L_TranslationPontM3.Safety_300.Idx318_EffectivePermitM3_Tremie := Translation.Safety.EffectivePermitM3_Tremie; // 🟢 Permis canonique vers Trémie
GVL_Troubleshooting.L_TranslationPontM3.Safety_300.Idx319_EffectivePermitM3_Maintenance := Translation.Safety.EffectivePermitM3_Maintenance; // 🟢 Permis canonique vers Maintenance/P1

GVL_Troubleshooting.L_TranslationPontM3.Control_400.Idx401_MotionAllowed := Translation.State.Ready;
GVL_Troubleshooting.L_TranslationPontM3.Control_400.Idx402_SetpointFreq_Hz := Translation.State.DriveFreqCmd_Hz;
GVL_Troubleshooting.L_TranslationPontM3.Control_400.Idx403_DriveControlWord := Translation.State.DriveControlWord;
GVL_Troubleshooting.L_TranslationPontM3.Control_400.Idx404_FinalInterlockState := Translation.State.FinalInterlockState;
GVL_Troubleshooting.L_TranslationPontM3.Control_400.Idx405_FinalInterlockReason := Translation.State.FinalInterlockReason;
GVL_Troubleshooting.L_TranslationPontM3.Control_400.Idx406_BrakeCommandOpenConfirmed := Translation.State.BrakeCommandOpenConfirmed;
GVL_Troubleshooting.L_TranslationPontM3.Control_400.Idx407_BrakeTimeoutElapsed := Translation.State.FinalBrakeTimeoutElapsed;

GVL_Troubleshooting.L_TranslationPontM3.Outputs_500.Idx501_CmdDriveControlWord := Translation.State.DriveControlWord;
GVL_Troubleshooting.L_TranslationPontM3.Outputs_500.Idx502_CmdDriveFreq_Hz := WORD_TO_UINT(CmdM3DriveFreqWord); // Consigne finale transmise, unité 0.01 Hz
GVL_Troubleshooting.L_TranslationPontM3.Outputs_500.Idx503_CmdBrakeRelease_RQ := Translation.State.BrakeCmd;

{endregion}

{region "§6 Diagnostic homing"}
// === 🎯 6. Diagnostic Chronologique Homing (HomingM1 & HomingM2) ===
// --- M1 ---
GVL_Troubleshooting.E_HomingM1.Step1_ModeAuthorized     := (Auth.Mode = E_Mode.MAINT_N1) OR (Auth.Mode = E_Mode.MAINT_N2);
GVL_Troubleshooting.E_HomingM1.Step2_WinchSelected      := (Auth.Mode <> E_Mode.MAINT_N2) OR (Auth.JoystickWinchSelectArbitrated = 1);
GVL_Troubleshooting.E_HomingM1.Step3_EncoderAvailable   := Network.EncoderM1.Operational AND NOT InputModuleFault;

GVL_Troubleshooting.E_HomingM1.HwIn_ContactorsReleased_DI := HwIn.Winch.M1_ContactorsReleased_DI;
GVL_Troubleshooting.E_HomingM1.HwIn_BrakeIsOpen_DI        := HwIn.Winch.M1_BrakeIsOpen_DI;
GVL_Troubleshooting.E_HomingM1.HwIn_TopPositionFree_DI    := HwIn.Winch.M1M2_TopPositionFree_DI;

GVL_Troubleshooting.E_HomingM1.Step4_ContactorsReleased := HwIn.Winch.M1_ContactorsReleased_DI;
GVL_Troubleshooting.E_HomingM1.Step5_BrakeApplied       := NOT HwIn.Winch.M1_BrakeIsOpen_DI;
GVL_Troubleshooting.E_HomingM1.TopPositionSensorActive  := Commun.TopPositionSensorActive;
GVL_Troubleshooting.E_HomingM1.BucketIsOpen             := WinchM2.Bucket.State.MechState.IsOpen;

GVL_Troubleshooting.E_HomingM1.AllConditionsMet := GVL_Troubleshooting.E_HomingM1.Step1_ModeAuthorized
                                              AND GVL_Troubleshooting.E_HomingM1.Step2_WinchSelected
                                              AND GVL_Troubleshooting.E_HomingM1.Step3_EncoderAvailable
                                              AND GVL_Troubleshooting.E_HomingM1.Step4_ContactorsReleased
                                              AND GVL_Troubleshooting.E_HomingM1.Step5_BrakeApplied;

GVL_Troubleshooting.E_HomingM1.HomingBusy      := WinchM1.State.Encoder.HomingBusy;
GVL_Troubleshooting.E_HomingM1.HomingDone      := WinchM1.State.Encoder.HomingDone;
GVL_Troubleshooting.E_HomingM1.HomingHomed     := WinchM1.State.Encoder.Homed;
GVL_Troubleshooting.E_HomingM1.HomingSuspect   := WinchM1.State.Encoder.HomingSuspect;
GVL_Troubleshooting.E_HomingM1.RejectErrorMask := WinchM1.State.Encoder.HomingErrorId;
GVL_Troubleshooting.E_HomingM1.TopContactLatched := MachineHoming.TopContactLatched;
GVL_Troubleshooting.E_HomingM1.TopContactCount   := MachineHoming.TopContactCount;

// --- M2 ---
GVL_Troubleshooting.F_HomingM2.Step1_ModeAuthorized     := (Auth.Mode = E_Mode.MAINT_N1) OR (Auth.Mode = E_Mode.MAINT_N2);
GVL_Troubleshooting.F_HomingM2.Step2_WinchSelected      := (Auth.Mode <> E_Mode.MAINT_N2) OR (Auth.JoystickWinchSelectArbitrated = 2);
GVL_Troubleshooting.F_HomingM2.Step3_EncoderAvailable   := Network.EncoderM2.Operational AND NOT InputModuleFault;

GVL_Troubleshooting.F_HomingM2.HwIn_ContactorsReleased_DI := HwIn.Winch.M2_ContactorsReleased_DI;
GVL_Troubleshooting.F_HomingM2.HwIn_BrakeIsOpen_DI        := HwIn.Winch.M2_BrakeIsOpen_DI;
GVL_Troubleshooting.F_HomingM2.HwIn_TopPositionFree_DI    := HwIn.Winch.M1M2_TopPositionFree_DI;

GVL_Troubleshooting.F_HomingM2.Step4_ContactorsReleased := HwIn.Winch.M2_ContactorsReleased_DI;
GVL_Troubleshooting.F_HomingM2.Step5_BrakeApplied       := NOT HwIn.Winch.M2_BrakeIsOpen_DI;
GVL_Troubleshooting.F_HomingM2.TopPositionSensorActive  := Commun.TopPositionSensorActive;
GVL_Troubleshooting.F_HomingM2.BucketIsOpen             := WinchM2.Bucket.State.MechState.IsOpen;

GVL_Troubleshooting.F_HomingM2.AllConditionsMet := GVL_Troubleshooting.F_HomingM2.Step1_ModeAuthorized
                                              AND GVL_Troubleshooting.F_HomingM2.Step2_WinchSelected
                                              AND GVL_Troubleshooting.F_HomingM2.Step3_EncoderAvailable
                                              AND GVL_Troubleshooting.F_HomingM2.Step4_ContactorsReleased
                                              AND GVL_Troubleshooting.F_HomingM2.Step5_BrakeApplied;

GVL_Troubleshooting.F_HomingM2.HomingBusy      := WinchM2.State.Encoder.HomingBusy;
GVL_Troubleshooting.F_HomingM2.HomingDone      := WinchM2.State.Encoder.HomingDone;
GVL_Troubleshooting.F_HomingM2.HomingHomed     := WinchM2.State.Encoder.Homed;
GVL_Troubleshooting.F_HomingM2.HomingSuspect   := WinchM2.State.Encoder.HomingSuspect;
GVL_Troubleshooting.F_HomingM2.RejectErrorMask := WinchM2.State.Encoder.HomingErrorId;
GVL_Troubleshooting.F_HomingM2.TopContactLatched := MachineHoming.TopContactLatched;
GVL_Troubleshooting.F_HomingM2.TopContactCount   := MachineHoming.TopContactCount;

{endregion}

{region "§7 Diagnostic chaine securite et AU"}
// === 🛡️ 7. Diagnostic Chronologique Chaîne de Sécurité & AU (Safety) ===
GVL_Troubleshooting.C_Safety.SimulationModeActive       := SimulationModeActive;
GVL_Troubleshooting.C_Safety.SimSafetyActive            := SimSafetyActive;

GVL_Troubleshooting.C_Safety.HwIn_EmergencyChainClosed_DI  := HwIn.Machine.EmergencyChainClosed_DI;
GVL_Troubleshooting.C_Safety.HwIn_PowerContactorEngaged_DI := HwIn.Machine.PowerContactorEngaged_DI;
GVL_Troubleshooting.C_Safety.HwIn_EmergencyBtnCut_HMI      := GVL_IHM.Emergency.Cmd.BtnEmergencyCutOff;

GVL_Troubleshooting.C_Safety.Step1_InputModulesOk       := NOT InputModuleFault;
GVL_Troubleshooting.C_Safety.Step2_EmergencyBtnNotCut   := NOT GVL_IHM.Emergency.Cmd.BtnEmergencyCutOff;
GVL_Troubleshooting.C_Safety.Step3_EmergencyChainClosed := HwIn.Machine.EmergencyChainClosed_DI;
GVL_Troubleshooting.C_Safety.Step4_ContactorReleased     := NOT HwIn.Machine.PowerContactorEngaged_DI;
GVL_Troubleshooting.C_Safety.Step5_ArmingAllowed        := EmergencyState.Armable;

GVL_Troubleshooting.C_Safety.ArmingStep            := EmergencyState.Step;
GVL_Troubleshooting.C_Safety.ArmingPulseActive    := ArmingPulseActive;
GVL_Troubleshooting.C_Safety.ArmingBusy           := EmergencyState.ArmingBusy;
GVL_Troubleshooting.C_Safety.LockoutActive        := EmergencyDiag.LockoutActive;
GVL_Troubleshooting.C_Safety.PowerContactorEngaged := HwIn.Machine.PowerContactorEngaged_DI;
GVL_Troubleshooting.C_Safety.PowerCutOffActive    := PowerCutOffActive;
GVL_Troubleshooting.C_Safety.PowerCutOffRequest   := Outputs.PowerCutOffRequest;
GVL_Troubleshooting.C_Safety.MaintainAActive      := MaintainAActive;
GVL_Troubleshooting.C_Safety.MaintainBActive      := MaintainBActive;

(* État final uniquement : ce n'est pas une précondition de réarmement. *)
GVL_Troubleshooting.C_Safety.AllConditionsMet := HwIn.Machine.EmergencyChainClosed_DI
                                            AND HwIn.Machine.PowerContactorEngaged_DI;
GVL_Troubleshooting.C_Safety.SafetyError          := EmergencyDiag.Error;
GVL_Troubleshooting.C_Safety.ArmingErrorId       := EmergencyDiag.ErrorId;
GVL_Troubleshooting.C_Safety.RedundancyTestFailed := EmergencyDiag.RedundancyTestFailed;
GVL_Troubleshooting.C_Safety.ArmingFailed         := EmergencyDiag.ArmFailed;
GVL_Troubleshooting.C_Safety.WasArmed             := EmergencyDiag.WasArmed;
GVL_Troubleshooting.C_Safety.LastAbortStep        := EmergencyDiag.LastAbortStep;
GVL_Troubleshooting.C_Safety.LastAbortCause       := EmergencyDiag.LastAbortCause;

{endregion}

{region "§8 Diagnostic CAN et joystick"}
// === 🕹️ 8. Diagnostic Chronologique Bus CAN & Joystick (Joystick) ===
GVL_Troubleshooting.D_Joystick.Step1_CanBusActive        := Network.BusCanOpen.Operational;
GVL_Troubleshooting.D_Joystick.Step2_JoystickOperational := Network.Joystick.Operational;
GVL_Troubleshooting.D_Joystick.HwIn_JoyBtnRaw_DI         := HwIn.Operator.JoyBtnRaw;
GVL_Troubleshooting.D_Joystick.NeutralXAct               := (HwIn.Operator.JoyXRaw_ANA1 >= 4800 AND HwIn.Operator.JoyXRaw_ANA1 <= 5200);
GVL_Troubleshooting.D_Joystick.NeutralYAct               := (HwIn.Operator.JoyYRaw_ANA2 >= 4800 AND HwIn.Operator.JoyYRaw_ANA2 <= 5200);
GVL_Troubleshooting.D_Joystick.Step3_DeadmanPressed      := HwIn.Operator.JoyBtnRaw;
GVL_Troubleshooting.D_Joystick.Step4_NeutralAcquired     := JoystickHMI.State.AtNeutral;
GVL_Troubleshooting.D_Joystick.DeadmanArmed             := JoystickHMI.State.DeadmanArmed;

GVL_Troubleshooting.D_Joystick.AllConditionsMet := GVL_Troubleshooting.D_Joystick.Step1_CanBusActive
                                              AND GVL_Troubleshooting.D_Joystick.Step2_JoystickOperational
                                              AND GVL_Troubleshooting.D_Joystick.DeadmanArmed;

GVL_Troubleshooting.D_Joystick.JoystickSelected := GVL_IHM.Modes.Cmd.TglJoystickMaster;
GVL_Troubleshooting.D_Joystick.SelJoystickWinch := GVL_IHM.Modes.Cmd.SelJoystickWinch;
GVL_Troubleshooting.D_Joystick.RawX             := HwIn.Operator.JoyXRaw_ANA1;
GVL_Troubleshooting.D_Joystick.RawY             := HwIn.Operator.JoyYRaw_ANA2;
GVL_Troubleshooting.D_Joystick.DeflectionX_Pct  := JoystickHMI.State.AxisCmdX.Deflection;
GVL_Troubleshooting.D_Joystick.DeflectionY_Pct  := JoystickHMI.State.AxisCmdY.Deflection;
// Direction exprimée en bits (ST_fbJoystick_AxisCmd) : conversion locale bits→INT (-1/0/+1),
// car ici on lit le struct (JoystickHMI.State.AxisCmdX/Y), pas le miroir FB DirectionX/Y.
IF JoystickHMI.State.AxisCmdX.DirectionPositive THEN
    GVL_Troubleshooting.D_Joystick.DirectionX := 1;
ELSIF JoystickHMI.State.AxisCmdX.DirectionNegative THEN
    GVL_Troubleshooting.D_Joystick.DirectionX := -1;
ELSE
    GVL_Troubleshooting.D_Joystick.DirectionX := 0;
END_IF;
IF JoystickHMI.State.AxisCmdY.DirectionPositive THEN
    GVL_Troubleshooting.D_Joystick.DirectionY := 1;
ELSIF JoystickHMI.State.AxisCmdY.DirectionNegative THEN
    GVL_Troubleshooting.D_Joystick.DirectionY := -1;
ELSE
    GVL_Troubleshooting.D_Joystick.DirectionY := 0;
END_IF;

{endregion}

{region "§9 Diagnostic mouvement treuil M1"}
// === ⚙️ 9. Diagnostic Chronologique Mouvement Treuil M1 (MotionM1) ===
GVL_Troubleshooting.N_MotionM1.Step1_PowerEngaged       := HwIn.Machine.PowerContactorEngaged_DI;
GVL_Troubleshooting.N_MotionM1.HwIn_PowerContactorEngaged_DI := HwIn.Machine.PowerContactorEngaged_DI;
GVL_Troubleshooting.N_MotionM1.HwIn_BrakeIsOpen_DI      := HwIn.Winch.M1_BrakeIsOpen_DI;
GVL_Troubleshooting.N_MotionM1.Cmd_BrakeRelease         := WinchM1.State.BrakeCmd;

GVL_Troubleshooting.N_MotionM1.Step2_ModeAuthorized     := (Auth.Mode <> E_Mode.DISABLE);
GVL_Troubleshooting.N_MotionM1.Step3_NotBusyOtherTask   := NOT WinchM1.State.Encoder.HomingBusy AND NOT (WinchM2.Bucket.State.FBState = E_State.BUSY);
GVL_Troubleshooting.N_MotionM1.Step4_MotionRequested    := WinchM1.State.Busy OR (WinchM1.State.SpeedCmd_Pct > 0.0);
GVL_Troubleshooting.N_MotionM1.RequestedDirection       := SEL(WinchM1.State.RelayFwd, SEL(WinchM1.State.RelayRev, 0, -1), 1);
GVL_Troubleshooting.N_MotionM1.RequestedSpeedPct        := WinchM1.State.SpeedCmd_Pct;
GVL_Troubleshooting.N_MotionM1.Step5_NoSafetyFault      := NOT WinchM1.Safety.SafeStop AND NOT WinchM1.Safety.ThermalFault;
GVL_Troubleshooting.N_MotionM1.Step6_DirectionAllowed   := SEL(GVL_Troubleshooting.N_MotionM1.RequestedDirection = 1, WinchM1.Safety.DescendPermit, WinchM1.Safety.AscentPermit);
GVL_Troubleshooting.N_MotionM1.Step7_BrakeReleased      := WinchM1.State.BrakeCmd AND WinchM1.State.BrakeCommandOpenConfirmed;
// 🛡️ T371 — honnêteté du diagnostic (M1). La barrière finale publie DÉJÀ son état et sa cause
// (FB_WinchOutputInterlock.st:54 State, :56 Reason), déjà routés jusqu'ici par
// FB_WinchStateProjection.st:112-115. L'ancien `NOT FinalInterlockError` ne lisait QUE le défaut
// bit0 (timeout confirmation frein, FB_WinchOutputInterlock.st:516-519 -> :528-532) : 4 refus
// RÉELS restaient affichés en vert — F1 RestartInhibit (:357-363), F2 ContactorStuckLatched
// (:364-373), F3 SafeStop/PermitFinalBlocked (:393-404, State laissé à READY et Reason à NONE),
// F4 RestartRequired/DeadTimePending (:424-429). On cesse de TRONQUER un état déjà publié.
// ⚠️ Latence N-1 assumée : WinchM1.State vient de la projection PRG_04_Treuils_Benne.st:1688-1696,
// qui lit l'instance de PRG_06_Outputs -> état daté d'un scan (~10 ms). USAGE DIAGNOSTIC UNIQUEMENT :
// aucune ligne de CONDUITE ne consomme Step8_InterlockState / Step8_InterlockReason.
// Le dernier terme (« demande moteur vivante SANS ordre de frein validé ») est le SEUL témoin publié
// qui distingue F3, où la barrière coupe les 6 ordres (:402-403) en laissant State = READY et Reason = NONE.
// 🔴 REX 2026-09-21 (revue indépendante T371, verdict BLOCK) : ce témoin NE DOIT SURTOUT PAS se
// construire sur `State.RelayFwd/RelayRev`. Ces champs viennent de FB_Winch
// (`FB_WinchStateProjection.st:102-103` <- `WinchM1Ref : FB_Winch`), c'est-à-dire de la DEMANDE —
// exactement le signal transmis à la barrière (`PRG_04_Treuils_Benne.st:1603-1604`
// `RequestedRelayFwd := instWinchM1.RelayFwd`). Comparer la demande à elle-même rend le terme
// TAUTOLOGIQUEMENT FAUX : `MotorRequest` implique déjà `RequestedRelayFwd XOR RequestedRelayRev`
// (`FB_WinchOutputInterlock.st:182`), donc F3 n'aurait JAMAIS été détecté et le test F3 aurait
// « passé » sur un état impossible en exploitation.
// ✅ Le seul témoin VALIDÉ publié est `State.BrakeCmd`, recopié de la SORTIE de la barrière
// (`FB_WinchStateProjection.st:108` <- `InterlockM1.BrakeCmd`, soit `RelayFwd OR RelayRev` VALIDÉS,
// `FB_WinchOutputInterlock.st:487`). Terme retenu : demande vivante ET aucun ordre validé.
// Recopie DIRECTE de l'énumération publiée (aucune projection, aucune conversion de type).
GVL_Troubleshooting.N_MotionM1.Step8_InterlockState  := WinchM1.State.FinalInterlockState;
GVL_Troubleshooting.N_MotionM1.Step8_InterlockReason := WinchM1.State.FinalInterlockReason;
GVL_Troubleshooting.N_MotionM1.Step8_OutputInterlockOk := NOT WinchM1.State.FinalInterlockError
                                                    AND NOT (WinchM1.State.FinalInterlockState = E_WinchFinalInterlockState.FAULT)
                                                    AND NOT (WinchM1.State.FinalInterlockState = E_WinchFinalInterlockState.DISABLED)
                                                    AND NOT (WinchM1.State.FinalInterlockState = E_WinchFinalInterlockState.WAIT_RESTART_DELAY)
                                                    AND NOT (WinchM1.State.FinalMotorRequest AND NOT WinchM1.State.BrakeCmd);

GVL_Troubleshooting.N_MotionM1.AllConditionsMet := GVL_Troubleshooting.N_MotionM1.Step1_PowerEngaged
                                              AND GVL_Troubleshooting.N_MotionM1.Step2_ModeAuthorized
                                              AND GVL_Troubleshooting.N_MotionM1.Step3_NotBusyOtherTask
                                              AND GVL_Troubleshooting.N_MotionM1.Step4_MotionRequested
                                              AND GVL_Troubleshooting.N_MotionM1.Step5_NoSafetyFault
                                              AND GVL_Troubleshooting.N_MotionM1.Step6_DirectionAllowed
                                              AND GVL_Troubleshooting.N_MotionM1.Step7_BrakeReleased
                                              AND GVL_Troubleshooting.N_MotionM1.Step8_OutputInterlockOk;

GVL_Troubleshooting.N_MotionM1.RelayFwdActive        := Outputs.M1RelayFwd;
GVL_Troubleshooting.N_MotionM1.RelayRevActive        := Outputs.M1RelayRev;
GVL_Troubleshooting.N_MotionM1.SpeedContactor1Active := Outputs.M1SpeedContactor1;

{endregion}

{region "§10 Diagnostic mouvement treuil M2"}
// === ⚙️ 10. Diagnostic Chronologique Mouvement Treuil M2 (MotionM2) ===
GVL_Troubleshooting.O_MotionM2.Step1_PowerEngaged       := HwIn.Machine.PowerContactorEngaged_DI;
GVL_Troubleshooting.O_MotionM2.HwIn_PowerContactorEngaged_DI := HwIn.Machine.PowerContactorEngaged_DI;
GVL_Troubleshooting.O_MotionM2.HwIn_BrakeIsOpen_DI      := HwIn.Winch.M2_BrakeIsOpen_DI;
GVL_Troubleshooting.O_MotionM2.Cmd_BrakeRelease         := WinchM2.State.BrakeCmd;

GVL_Troubleshooting.O_MotionM2.Step2_ModeAuthorized     := (Auth.Mode <> E_Mode.DISABLE);
GVL_Troubleshooting.O_MotionM2.Step3_NotBusyOtherTask   := NOT WinchM2.State.Encoder.HomingBusy;
GVL_Troubleshooting.O_MotionM2.Step4_MotionRequested    := WinchM2.State.Busy OR (WinchM2.State.SpeedCmd_Pct > 0.0);
GVL_Troubleshooting.O_MotionM2.RequestedDirection       := SEL(WinchM2.State.RelayFwd, SEL(WinchM2.State.RelayRev, 0, -1), 1);
GVL_Troubleshooting.O_MotionM2.RequestedSpeedPct        := WinchM2.State.SpeedCmd_Pct;
GVL_Troubleshooting.O_MotionM2.Step5_NoSafetyFault      := NOT WinchM2.Safety.SafeStop AND NOT WinchM2.Safety.ThermalFault AND NOT WinchM2.Safety.SlackCable;
GVL_Troubleshooting.O_MotionM2.Step6_DirectionAllowed   := SEL(GVL_Troubleshooting.O_MotionM2.RequestedDirection = 1, WinchM2.Safety.DescendPermit, WinchM2.Safety.AscentPermit);
GVL_Troubleshooting.O_MotionM2.Step7_BrakeReleased      := WinchM2.State.BrakeCmd AND WinchM2.State.BrakeCommandOpenConfirmed;
// 🛡️ T371 — honnêteté du diagnostic (M2), même patron que M1 ci-dessus (source :
// FB_WinchStateProjection.st:179-182, barrière FB_WinchOutputInterlock.st:54/:56, refus F1-F4
// aux sites :357-363 / :364-373 / :393-404 / :424-429). Lecture N-1, DIAGNOSTIC UNIQUEMENT.
// Idem M1 : le témoin F3 est `BrakeCmd` (SORTIE validée, projection :175) et JAMAIS les relais
// `RelayFwd/RelayRev` de la demande (tautologie — REX revue T371 du 2026-09-21).
GVL_Troubleshooting.O_MotionM2.Step8_InterlockState  := WinchM2.State.FinalInterlockState;
GVL_Troubleshooting.O_MotionM2.Step8_InterlockReason := WinchM2.State.FinalInterlockReason;
GVL_Troubleshooting.O_MotionM2.Step8_OutputInterlockOk := NOT WinchM2.State.FinalInterlockError
                                                    AND NOT (WinchM2.State.FinalInterlockState = E_WinchFinalInterlockState.FAULT)
                                                    AND NOT (WinchM2.State.FinalInterlockState = E_WinchFinalInterlockState.DISABLED)
                                                    AND NOT (WinchM2.State.FinalInterlockState = E_WinchFinalInterlockState.WAIT_RESTART_DELAY)
                                                    AND NOT (WinchM2.State.FinalMotorRequest AND NOT WinchM2.State.BrakeCmd);

GVL_Troubleshooting.O_MotionM2.AllConditionsMet := GVL_Troubleshooting.O_MotionM2.Step1_PowerEngaged
                                              AND GVL_Troubleshooting.O_MotionM2.Step2_ModeAuthorized
                                              AND GVL_Troubleshooting.O_MotionM2.Step3_NotBusyOtherTask
                                              AND GVL_Troubleshooting.O_MotionM2.Step4_MotionRequested
                                              AND GVL_Troubleshooting.O_MotionM2.Step5_NoSafetyFault
                                              AND GVL_Troubleshooting.O_MotionM2.Step6_DirectionAllowed
                                              AND GVL_Troubleshooting.O_MotionM2.Step7_BrakeReleased
                                              AND GVL_Troubleshooting.O_MotionM2.Step8_OutputInterlockOk;

GVL_Troubleshooting.O_MotionM2.RelayFwdActive        := Outputs.M2RelayFwd;
GVL_Troubleshooting.O_MotionM2.RelayRevActive        := Outputs.M2RelayRev;
GVL_Troubleshooting.O_MotionM2.SpeedContactor1Active := Outputs.M2SpeedContactor1;

{endregion}

{region "§11 Diagnostic mouvement translation M3"}
// === ⚙️ 10bis. Diagnostic Chronologique Mouvement Translation M3 (MotionM3) ===
GVL_Troubleshooting.P_MotionM3.Step1_PowerEngaged       := HwIn.Machine.PowerContactorEngaged_DI;
GVL_Troubleshooting.P_MotionM3.HwIn_PowerContactorEngaged_DI := HwIn.Machine.PowerContactorEngaged_DI;
GVL_Troubleshooting.P_MotionM3.HwIn_BrakeIsOpen_DI      := HwIn.Translation.M3_BrakeIsOpen_DI;
GVL_Troubleshooting.P_MotionM3.Cmd_BrakeRelease         := Translation.State.BrakeCmd;

GVL_Troubleshooting.P_MotionM3.Step2_ModeAuthorized     := (Auth.Mode <> E_Mode.DISABLE);
GVL_Troubleshooting.P_MotionM3.Step3_NotBusyOtherTask   := TRUE; // Aucune tâche exclusive connue bloquant M3 (pas de homing translation)
GVL_Troubleshooting.P_MotionM3.Step4_MotionRequested    := Translation.State.Busy OR (Translation.State.SpeedCmd_Pct > 0.0);
// Conversion locale uniquement pour compatibilité de l'index diagnostic historique :
// les contrats M3 et les commandes utilisent les deux bits explicites.
GVL_Troubleshooting.P_MotionM3.RequestedDirection       := SEL(Translation.State.ActiveTremie,
                                                               SEL(Translation.State.ActiveMaintenance, -1, 0), 1);
GVL_Troubleshooting.P_MotionM3.RequestedSpeedPct        := Translation.State.SpeedCmd_Pct;
GVL_Troubleshooting.P_MotionM3.Step5_NoSafetyFault      := NOT Translation.Safety.SafeStop AND NOT Translation.State.Error;
GVL_Troubleshooting.P_MotionM3.Step6_DirectionAllowed   := SEL(GVL_Troubleshooting.P_MotionM3.RequestedDirection = 1, Translation.Safety.EffectivePermitM3_Maintenance, Translation.Safety.EffectivePermitM3_Tremie); // Permis canoniques M3 — HeightInterlockBlocking reste un blocage séparé
GVL_Troubleshooting.P_MotionM3.Step7_BrakeReleased      := Translation.State.BrakeCmd AND Translation.State.BrakeCommandOpenConfirmed;
// 🛡️ T371 — axe M3 : état et cause publiés, décision inchangée sur le seul témoin ACTIF disponible.
// Pourquoi pas plus ici : (1) la barrière finale M3 ne publie AUCUN état machine — PRG_05_Translation.st:749-755
// dérive FinalInterlockState de Fault.Error seul (READY/ERROR), et ses ordres validés (DriveControlWord,
// DriveFreqCmd) ne sont PAS publiés vers l'IHM (TranslationState.DriveControlWord :717 recopie la DEMANDE
// de FB_Translation, pas l'ordre validé de la barrière) -> aucun témoin « ordre réellement délivré » ;
// (2) `FinalInterlockReason` est MÉMORISÉ et n'est JAMAIS remis à NONE après acquittement
// (FB_TranslationOutputInterlock.st:123-130 lève RestartInhibit sans toucher Reason ; seul le gate :80
// le remet à NONE) -> l'utiliser dans la décision créerait un faux ROUGE PERMANENT après un acquittement.
// Il est donc PUBLIÉ pour le technicien, sans servir de preuve de refus actif.
// Le rapprochement avec la vérité Control_400 (Idx404/Idx405) devient ainsi lisible dans la checklist.
// M3 ne publie qu'un état DÉRIVÉ du défaut (PRG_05:751-755) : projection EXPLICITE sur le vocabulaire
// commun du DUT (E_State.READY -> READY, E_State.ERROR -> FAULT) — aucune donnée inventée, aucune
// conversion de type. Les 3 raisons M3 sont identiques à celles de la famille commune.
IF Translation.State.FinalInterlockState = E_State.ERROR THEN
    GVL_Troubleshooting.P_MotionM3.Step8_InterlockState := E_WinchFinalInterlockState.FAULT;
ELSE
    GVL_Troubleshooting.P_MotionM3.Step8_InterlockState := E_WinchFinalInterlockState.READY;
END_IF;
IF Translation.State.FinalInterlockReason = E_TranslationFinalInterlockReason.RESTART_INHIBITED THEN
    GVL_Troubleshooting.P_MotionM3.Step8_InterlockReason := E_WinchFinalInterlockReason.RESTART_INHIBITED;
ELSIF Translation.State.FinalInterlockReason = E_TranslationFinalInterlockReason.BRAKE_COMMAND_NOT_CONFIRMED THEN
    GVL_Troubleshooting.P_MotionM3.Step8_InterlockReason := E_WinchFinalInterlockReason.BRAKE_COMMAND_NOT_CONFIRMED;
ELSE
    GVL_Troubleshooting.P_MotionM3.Step8_InterlockReason := E_WinchFinalInterlockReason.NONE;
END_IF;
GVL_Troubleshooting.P_MotionM3.Step8_OutputInterlockOk := NOT Translation.State.FinalInterlockError
                                                    AND NOT (Translation.State.FinalInterlockState = E_State.ERROR);

GVL_Troubleshooting.P_MotionM3.AllConditionsMet := GVL_Troubleshooting.P_MotionM3.Step1_PowerEngaged
                                              AND GVL_Troubleshooting.P_MotionM3.Step2_ModeAuthorized
                                              AND GVL_Troubleshooting.P_MotionM3.Step3_NotBusyOtherTask
                                              AND GVL_Troubleshooting.P_MotionM3.Step4_MotionRequested
                                              AND GVL_Troubleshooting.P_MotionM3.Step5_NoSafetyFault
                                              AND GVL_Troubleshooting.P_MotionM3.Step6_DirectionAllowed
                                              AND GVL_Troubleshooting.P_MotionM3.Step7_BrakeReleased
                                              AND GVL_Troubleshooting.P_MotionM3.Step8_OutputInterlockOk;

// 🔌 M3 piloté par variateur AC600 (pas de relais/contacteur de palier comme M1/M2) : ces
// champs restent des indicateurs de sens actif, pas des retours relais physiques réels.
GVL_Troubleshooting.P_MotionM3.RelayFwdActive        := Translation.State.ActiveTremie AND Translation.State.Busy;
GVL_Troubleshooting.P_MotionM3.RelayRevActive        := Translation.State.ActiveMaintenance AND Translation.State.Busy;
GVL_Troubleshooting.P_MotionM3.SpeedContactor1Active := FALSE; // Non applicable — M3 n'a pas de contacteur de vitesse par palier

{endregion}

{region "§12 Images entrees reelles et simulees"}
// === 📥 11. Image Complète des Entrées Réelles / Simulées (Inputs) ===
GVL_Troubleshooting.B_Inputs := HwIn;
{endregion}

{region "§13 Séquenceur de cycle semi-automatique"}
// === 🔄 12. Diagnostic Chronologique Séquenceur Semi-Auto (CycleSemiAuto) ===
GVL_Troubleshooting.G_CycleSemiAuto.Idx101_ModeSemiAutoActive        := (Auth.Mode = E_Mode.SEMI_AUTO);
GVL_Troubleshooting.G_CycleSemiAuto.Idx102_PowerAndSafetyOk          := HwIn.Machine.PowerContactorEngaged_DI;
GVL_Troubleshooting.G_CycleSemiAuto.Idx103_HeartbeatIhmOk            := Commun.HeartbeatIhmOk;
GVL_Troubleshooting.G_CycleSemiAuto.Idx104_DeadmanArmed              := JoystickDeadmanArmed;
GVL_Troubleshooting.G_CycleSemiAuto.Idx105_MancheDeflechi            := NOT JoystickAtNeutral;
GVL_Troubleshooting.G_CycleSemiAuto.Idx106_HomedM1M2                 := HomedM1 AND HomedM2;
GVL_Troubleshooting.G_CycleSemiAuto.Idx107_StartCycleRequest         := CycleStartRequest;
GVL_Troubleshooting.G_CycleSemiAuto.Idx108_AbortCycleRequest         := CycleAbortRequest;

GVL_Troubleshooting.G_CycleSemiAuto.Idx201_Ready                     := CycleReady;
GVL_Troubleshooting.G_CycleSemiAuto.Idx202_Busy                      := CycleAutoBusy;
GVL_Troubleshooting.G_CycleSemiAuto.Idx203_Done                      := CycleDone;
GVL_Troubleshooting.G_CycleSemiAuto.Idx204_Error                     := CycleError;
GVL_Troubleshooting.G_CycleSemiAuto.Idx205_ErrorId                   := CycleErrorId;
GVL_Troubleshooting.G_CycleSemiAuto.Idx217_FaultLatched               := CycleFaultLatched;
GVL_Troubleshooting.G_CycleSemiAuto.Idx218_FaultLatchedId             := CycleFaultLatchedId;
GVL_Troubleshooting.G_CycleSemiAuto.Idx219_CycleChecksInhibited       := CycleChecksInhibited;
GVL_Troubleshooting.G_CycleSemiAuto.Idx220_IgnoredCycleCheckId        := CycleIgnoredCheckId;
GVL_Troubleshooting.G_CycleSemiAuto.Idx222_ForceStepResult            := CycleForceStepResult;
GVL_Troubleshooting.G_CycleSemiAuto.Idx206_Step                      := CycleStep;
GVL_Troubleshooting.G_CycleSemiAuto.Idx207_StepStr                   := CycleStepStr;
GVL_Troubleshooting.G_CycleSemiAuto.Idx208_StepAtError               := CycleStepAtError;
GVL_Troubleshooting.G_CycleSemiAuto.Idx209_WaitingForOperator        := CycleWaitingForOperator;
GVL_Troubleshooting.G_CycleSemiAuto.Idx210_WaitingForProcess         := CycleWaitingForProcess;
GVL_Troubleshooting.G_CycleSemiAuto.Idx211_OperatorActionId          := CycleOperatorActionId;
GVL_Troubleshooting.G_CycleSemiAuto.Idx212_OperatorAction            := CycleOperatorAction;
GVL_Troubleshooting.G_CycleSemiAuto.Idx213_ExpectedAxis              := CycleExpectedAxis;
GVL_Troubleshooting.G_CycleSemiAuto.Idx214_ExpectedDirection         := CycleExpectedDirection;
GVL_Troubleshooting.G_CycleSemiAuto.Idx215_WaitingResume             := (Auth.Mode <> E_Mode.SEMI_AUTO) AND (CycleStep <> E_AutoCycleStep.AX0_REPOS) AND (CycleStep <> E_AutoCycleStep.AX18_DONE_SYNC) AND (CycleStep <> E_AutoCycleStep.AX_STAB);
GVL_Troubleshooting.G_CycleSemiAuto.Idx216_PausedState               := CycleStep;

GVL_Troubleshooting.G_CycleSemiAuto.Idx301_TargetPosition            := CycleTargetPosition;
GVL_Troubleshooting.G_CycleSemiAuto.Idx302_TargetDepth_M             := CycleTargetDepth_M;
GVL_Troubleshooting.G_CycleSemiAuto.Idx303_KoboldBottomTouch         := CycleKoboldBottomTouch;
GVL_Troubleshooting.G_CycleSemiAuto.Idx304_SpeedMismatchActive       := CycleSpeedMismatchActive;
GVL_Troubleshooting.G_CycleSemiAuto.Idx305_LimitLegalReached         := CycleLimitLegalReached;
GVL_Troubleshooting.G_CycleSemiAuto.Idx306_WinchSyncError            := CycleWinchSyncError;
GVL_Troubleshooting.G_CycleSemiAuto.Idx307_M1SpeedStepApplied        := CycleM1SpeedStepApplied;
GVL_Troubleshooting.G_CycleSemiAuto.Idx308_M2SpeedStepApplied        := CycleM2SpeedStepApplied;
GVL_Troubleshooting.G_CycleSemiAuto.Idx309_AutoDiveM2Step5Active     := CycleAutoDiveM2Step5Active;
GVL_Troubleshooting.G_CycleSemiAuto.Idx310_M1SpeedStepAtFault        := CycleM1SpeedStepAtFault;
GVL_Troubleshooting.G_CycleSemiAuto.Idx311_M2SpeedStepAtFault        := CycleM2SpeedStepAtFault;
{endregion}

{region "§14 Trace de blocage terrain (winch M1/M2 + translation M3)"}
// === 🕵️ 13. Trace de blocage terrain (ST_TraceWinch / ST_TraceTranslation) ===
// Pur recopie des traces publiées par PRG_04 (§8bis) et PRG_05 (§4bis). Aucun calcul métier ici.
GVL_Troubleshooting.Q_TraceWinchM1     := WinchM1Trace;
GVL_Troubleshooting.R_TraceWinchM2     := WinchM2Trace;
GVL_Troubleshooting.S_TraceTranslation := TranslationTrace;
GVL_Troubleshooting.T_Permits           := Permits;
{endregion}
